(* PLC project FB_BackwashGraph, s7-to-codesys s7conv 1.2.0 *)
(* stored: creationDateTime 2026-10-20T00:00:00 *)

FUNCTION_BLOCK FB_BackwashGraph_Sfc
  VAR_INPUT
    SFCInit : BOOL;  (* INIT_SQ: начальное состояние (флаг SFC) *)
    xStart : BOOL;  (* Пуск промывки *)
    xLevelLow : BOOL;  (* Уровень ниже сливного *)
    xLevelHigh : BOOL;  (* Фильтр заполнен *)
    xShortWash : BOOL;  (* Короткая промывка (без продувки) *)
    xPumpOk : BOOL := TRUE;  (* Насос промывки исправен *)
    xValveFault : BOOL;  (* Неисправность сливной задвижки *)
    Drain_SvErr : BOOL;  (* шаг S2: ошибка контроля (защёлка обёртки) *)
  END_VAR
  VAR_OUTPUT
    xIdle_N1 : BOOL;  (* шаг S1: действие N *)
    xDrain_N1 : BOOL;  (* шаг S2: действие N *)
    xDrain_S2 : BOOL;  (* шаг S2: действие N *)
    xDrain_P3 : BOOL;  (* шаг S2: действие P *)
    xDrain_Active : BOOL;  (* шаг S2: действие N *)
    xAir_N1 : BOOL;  (* шаг S3: действие N *)
    xAir_D2 : BOOL;  (* шаг S3: действие D *)
    xRinse_N1 : BOOL;  (* шаг S4: действие N *)
    xQuickRinse_N1 : BOOL;  (* шаг S5: действие N *)
    xRefill_N1 : BOOL;  (* шаг S6: действие N *)
    xRefill_R2 : BOOL;  (* шаг S6: действие N *)
  END_VAR

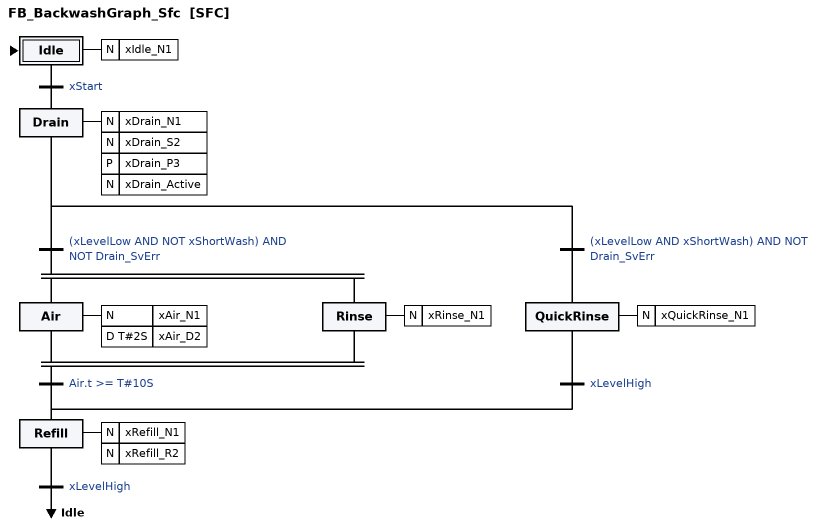
INITIAL_STEP Idle:
  xIdle_N1(N);
END_STEP
TRANSITION FROM Idle TO Drain
  := xStart;
END_TRANSITION
STEP Drain:
  xDrain_N1(N);
  xDrain_S2(N);
  xDrain_P3(P);
  xDrain_Active(N);
END_STEP
TRANSITION FROM Drain TO (Air, Rinse)
  := (xLevelLow AND NOT xShortWash) AND NOT Drain_SvErr;
END_TRANSITION
TRANSITION FROM Drain TO QuickRinse
  := (xLevelLow AND xShortWash) AND NOT Drain_SvErr;
END_TRANSITION
STEP Air:
  xAir_N1(N);
  xAir_D2(D, T#2S);
END_STEP
TRANSITION FROM (Air, Rinse) TO Refill
  := Air.t >= T#10S;
END_TRANSITION
STEP Rinse:
  xRinse_N1(N);
END_STEP
STEP QuickRinse:
  xQuickRinse_N1(N);
END_STEP
TRANSITION FROM QuickRinse TO Refill
  := xLevelHigh;
END_TRANSITION
STEP Refill:
  xRefill_N1(N);
  xRefill_R2(N);
END_STEP
TRANSITION FROM Refill TO Idle
  := xLevelHigh;
END_TRANSITION
END_FUNCTION_BLOCK

FUNCTION_BLOCK FB_BackwashGraph
  VAR_INPUT
    OFF_SQ : BOOL;  (* Выключить последовательность *)
    INIT_SQ : BOOL;  (* Начальное состояние *)
    ACK_EF : BOOL;  (* Квитирование ошибок контроля *)
    xStart : BOOL;  (* Пуск промывки *)
    xLevelLow : BOOL;  (* Уровень ниже сливного *)
    xLevelHigh : BOOL;  (* Фильтр заполнен *)
    xShortWash : BOOL;  (* Короткая промывка (без продувки) *)
    xPumpOk : BOOL := TRUE;  (* Насос промывки исправен *)
    xValveFault : BOOL;  (* Неисправность сливной задвижки *)
  END_VAR
  VAR_OUTPUT
    ERR_FLT : BOOL;  (* Ошибка контроля (до квитирования) *)
    xReady : BOOL;  (* Готов к промывке *)
    xDrainValve : BOOL;  (* Сливная задвижка *)
    xBlower : BOOL;  (* Воздуходувка *)
    xAirValve : BOOL;  (* Задвижка воздуха *)
    xWashPump : BOOL;  (* Насос промывки *)
    xInletValve : BOOL;  (* Задвижка подачи *)
    xWashActive : BOOL;  (* Промывка идёт *)
    xValvesBusy : BOOL;  (* Задвижки в работе *)
    iWashCount : INT;  (* Число промывок *)
  END_VAR
  VAR
    fbSfc : FB_BackwashGraph_Sfc;  (* последовательность SFC *)
    Drain_SvErr : BOOL;  (* шаг S2: ошибка контроля *)
  END_VAR

// Сгенерировано s7conv из samples/lang/FB_BackwashGraph.xml (S7-GRAPH, стратегия sfc):
// SFC FB_BackwashGraph_Sfc и обёртка FB_BackwashGraph с интерфейсом блока GRAPH.
// Квитирование ошибок контроля (ACK_EF) и INIT_SQ — до вызова SFC: в этом цикле переход возможен
IF ACK_EF OR INIT_SQ THEN
    Drain_SvErr := FALSE;
END_IF
fbSfc(SFCInit := INIT_SQ, xStart := xStart, xLevelLow := xLevelLow, xLevelHigh := xLevelHigh,
      xShortWash := xShortWash, xPumpOk := xPumpOk, xValveFault := xValveFault, Drain_SvErr := Drain_SvErr);
// Действия GRAPH по флагам IEC-действий SFC
xReady := (fbSfc.xIdle_N1 OR INIT_SQ);
xDrainValve := (fbSfc.xDrain_N1 AND NOT INIT_SQ);
xBlower := (fbSfc.xAir_N1 AND NOT INIT_SQ);
xAirValve := (fbSfc.xAir_D2 AND NOT INIT_SQ);
xWashPump := (fbSfc.xRinse_N1 AND NOT INIT_SQ) AND (xPumpOk) OR (fbSfc.xQuickRinse_N1 AND NOT INIT_SQ);
xInletValve := (fbSfc.xRefill_N1 AND NOT INIT_SQ);
IF (fbSfc.xDrain_S2 AND NOT INIT_SQ) THEN // S2: S xWashActive
    xWashActive := TRUE;
END_IF
IF (fbSfc.xDrain_P3 AND NOT INIT_SQ) THEN // S2: событие S1
    iWashCount := iWashCount + 1;
END_IF
IF (fbSfc.xRefill_R2 AND NOT INIT_SQ) THEN // S6: R xWashActive
    xWashActive := FALSE;
END_IF
// Контроль шагов: ошибка защёлкивается до ACK_EF
IF (fbSfc.xDrain_Active AND NOT INIT_SQ) AND (xValveFault) THEN
    Drain_SvErr := TRUE;
END_IF
ERR_FLT := Drain_SvErr;
// Постоперация 1
xValvesBusy := xDrainValve OR xInletValve;
END_FUNCTION_BLOCK
